FUNCTION_BLOCK FB_Emergency_Shutdown
VAR_INPUT
END_VAR
VAR_OUTPUT
	bTrip : BOOL;          // TRUE = systemet skal stoppes
END_VAR
VAR_IN_OUT
	Motor_ON_OFF      : BOOL;
	bControllerActive : BOOL;
	Motor_speed       : INT;
	Gas_Valve         : INT;
	Flow_Valve_1      : INT;
	Level_Valve_1     : INT;
	Level_Valve_2     : INT;
	Level_Valve_3     : INT;
END_VAR

//MAIN . fbPressAlarm . bAlarm
 //│          │           │
// │          │           └─ variabelen bAlarm inne i den blokken
// │          └─ instansen fbPressAlarm, som er deklarert i MAIN
// └─ programmet MAIN

//Instans: typen er en funksjonsblokk. Den holder en hel pakke, med innganger, utganger og internt minne, og den har kode som kan kjøres.

// Gas_Valve := REAL_TO_INT(262.14 * Prosent + 6553);

// Setter maskinen i safe state
VAR
	fbTripLatch: SR;
END_VAR
VAR // added by the converter: edge detectors and wires of the graphical bodies
    _w1 : BOOL;
END_VAR

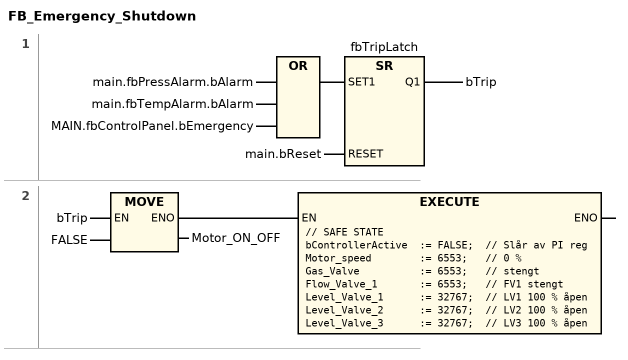
// NETWORK 1
fbTripLatch(SET1 := main.fbPressAlarm.bAlarm OR main.fbTempAlarm.bAlarm OR MAIN.fbControlPanel.bEmergency, RESET := main.bReset); // SR
bTrip := fbTripLatch.Q1;

// NETWORK 2
_w1 := bTrip;
IF _w1 THEN Motor_ON_OFF := FALSE; END_IF
IF _w1 THEN
    // SAFE STATE
    bControllerActive  := FALSE;  // Slår av PI reg 
    Motor_speed        := 6553;   // 0 %
    Gas_Valve          := 6553;   // stengt
    Flow_Valve_1       := 6553;   // FV1 stengt
    Level_Valve_1      := 32767;  // LV1 100 % åpen
    Level_Valve_2      := 32767;  // LV2 100 % åpen
    Level_Valve_3      := 32767;  // LV3 100 % åpen
END_IF

END_FUNCTION_BLOCK

(* stored: Version 1.1.0.1, ProductVersion 3.1.4026.21
   POU FB_Emergency_Shutdown: Id {70ab5e32-1960-4844-8ef8-2f5ee2dcfeef}, SpecialFunc None *)
